{attribute 'qualified_only'}
{attribute 'strict'}
{attribute 'to_string'}
TYPE E_Lint :
(
	eOptionA := 0,
	eOptionB,
	eOptionC
) LINT;
END_TYPE

(* stored: Version 1.1.0.1, ProductVersion 3.1.4026.19
   DUT E_Lint: Id {dbdfab39-b5c4-43d2-80a6-3102a8d14bec} *)
